Fanuc KAREL source: KD00054.KL

PROGRAM KD00054
%NOLOCKGROUP
VAR
  I: INTEGER
  J: INTEGER
  B: BOOLEAN
  R: REAL
  S: STRING[80]
BEGIN
  CONDITION[1]:
  WHEN DIN[1] = ON DO
    I = 7
  ENDCONDITION
END KD00054
